SUBAPPLICATION Uebung_OPC_L07_AX (* Wie Training_07 (Adapter-Variante von 05), lokal: Set/Reset per localhost, Zustand lokal per PUBLISH *)
  (* Standard: 61499-2; Description: Copyright (c) 2026 Meisterschulen am Ostbahnhof This program and the accompanying materials are made available under the terms of the Eclipse Public License 2.0 which is available at https://www.eclipse.org/legal/epl-2.0/ SPDX-License-Identifier: EPL-2.0 *)
  (* Version 1.0, 2026-10-18, Franz Höpfinger, Meisterschulen am Ostbahnhof, Aus SubApp_PC_A + SubApp_PC_B von test_VV zusammengefuehrt, lokale Varianten der Bausteine *)
  PACKAGE Meins::OPC_UA_Lokal;
  IMPORT Uebungen::const::UT::DefaultPool::SoftKey_F1;
  IMPORT Uebungen::const::UT::DefaultPool::SoftKey_F2;
  IMPORT Meins::OPC_UA_Lokal::const::OpcUaLokal::SR2_SET_CALL;
  IMPORT Meins::OPC_UA_Lokal::const::OpcUaLokal::SR2_RESET_CALL;
  IMPORT Meins::OPC_UA_Lokal::const::OpcUaLokal::SR2_STATE_READ;
  IMPORT logiBUS::io::DQ::logiBUS_DO::Output_Q1;
  IMPORT Meins::OPC_UA_Lokal::const::OpcUaLokal::SR2_SET_METHOD;
  IMPORT Meins::OPC_UA_Lokal::const::OpcUaLokal::SR2_RESET_METHOD;
  IMPORT Meins::OPC_UA_Lokal::const::OpcUaLokal::SR2_STATE_WRITE;
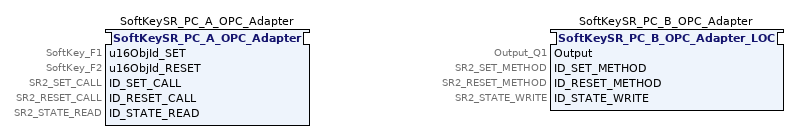
  SUBAPPS
    SoftKeySR_PC_A_OPC_Adapter : MyLib::sys::SoftKeySR_PC_A_OPC_Adapter(u16ObjId_SET := SoftKey_F1, u16ObjId_RESET := SoftKey_F2, ID_SET_CALL := SR2_SET_CALL, ID_RESET_CALL := SR2_RESET_CALL, ID_STATE_READ := SR2_STATE_READ);
    SoftKeySR_PC_B_OPC_Adapter : MyLib::sys::SoftKeySR_PC_B_OPC_Adapter_LOC(Output := Output_Q1, ID_SET_METHOD := SR2_SET_METHOD, ID_RESET_METHOD := SR2_RESET_METHOD, ID_STATE_WRITE := SR2_STATE_WRITE);
  END_SUBAPPS
END_SUBAPPLICATION
